(* IEC 61131-3 sources: plc-workbench/experiments/general_tasks_r6/followup/restart_delay, 2 files *)

(* ---- candidate_01.st ---- *)
FUNCTION_BLOCK RestartDelay
VAR_INPUT
    request : BOOL;
    inhibit : BOOL;
    delay : TIME;
END_VAR
VAR_OUTPUT
    running : BOOL;
END_VAR
VAR
    timer : TON;
END_VAR

timer(IN := request AND NOT inhibit, PT := delay);
running := timer.Q;

END_FUNCTION_BLOCK

(* ---- candidate_final.st ---- *)
FUNCTION_BLOCK RestartDelay
VAR_INPUT
    request : BOOL;
    inhibit : BOOL;
    delay : TIME;
END_VAR
VAR_OUTPUT
    running : BOOL;
END_VAR
VAR
    timer : TON;
END_VAR

timer(IN := request AND NOT inhibit, PT := delay);
running := timer.Q;

END_FUNCTION_BLOCK
